TYPE ST_KUKA_REF : FB_KUKA_REF;
END_TYPE

(* stored: Version 1.1.0.1, ProductVersion 3.1.4024.15
   DUT ST_KUKA_REF: Id {0f4980ae-8cf9-44fc-b254-92b6468a9fcc} *)
